(* PLC project Tank, plca e2e 1 *)
(* stored: creationDateTime 2026-10-25T10:00:00, modificationDateTime 2026-10-25T10:00:00 *)

PROGRAM TankCheck
  VAR
    rVolume : REAL;
    bFull : BOOL;
  END_VAR

bFull := rVolume = 100.0;
END_PROGRAM
